INTERFACE I_MoverDetectionAlgorithm EXTENDS i_Task


METHOD Abort : HRESULT
VAR_INPUT
END_VAR
END_METHOD

PROPERTY DetectedMoverCount : UDINT
GET
END_GET
END_PROPERTY

METHOD Reset : HRESULT
VAR_INPUT
END_VAR
END_METHOD

METHOD SetComponents : BOOL
VAR_INPUT
	XtsTracks : ARRAY[0..TcIoXtsEnvironmentParameterList.MaxXtsTracksPerXpu] OF I_XtsTrack;
	MoverArray : ARRAY[0..TcIoXtsEnvironmentParameterList.MaxXtsMoversPerXpu] OF I_XtsMover;
	XPU : I_TcIoXtsProcessingUnit;
END_VAR
END_METHOD

METHOD Start : HRESULT
VAR_INPUT
END_VAR
END_METHOD

END_INTERFACE

(* stored: Version 1.1.0.1
   Itf I_MoverDetectionAlgorithm: Id {33d5f92a-ed58-4708-a470-1691ea7312ec}
   Method Abort: Id {dd31e5d6-eaa0-46fc-b5ea-c32a606fe694}
   Property DetectedMoverCount: Id {56fda154-0eef-4840-bd70-7005b92b3e2c}
   Get Get: Id {920f32c2-a114-4e59-b985-4870f90b8bff}
   Method Reset: Id {b7d11555-81bd-4227-a0a5-39d83d020680}
   Method SetComponents: Id {a706bd72-b2c6-4d16-b576-edfdb2cd5c7a}
   Method Start: Id {b150b5fa-d8d3-410a-8834-e2b67794974e} *)
